DATA_BLOCK "naut_SfcFinalScan_DB"
{ S7_Optimized_Access := 'TRUE' }
VERSION : 0.1
"naut_SfcFinalScan"

BEGIN

END_DATA_BLOCK
